Yaskawa INFORM job: -DEFRO-70-PRZYLACZE-70-NOWE.JBI

/JOB
//NAME -DEFRO-70-PRZYLACZE-70-NOWE
//POS
///NPOS 61,61,61,0,0,0
///TOOL 0
///POSTYPE PULSE
///PULSE
C00000=-281,-101163,-84214,3730,-80188,-1936
C00001=-283,-101162,-84213,3710,-80188,-1936
C00002=116617,-39062,-41553,1138,-40446,20
C00003=97332,10008,-65831,-77395,-56626,78097
C00004=97332,10036,-65835,-77406,-56622,78106
C00005=126597,-12792,-74683,9116,-14112,37031
C00006=129578,-9389,-72169,26197,-17561,29790
C00007=143171,23000,-49885,51799,-48783,19450
C00008=142289,27625,-43624,46606,-52109,19593
C00009=140707,34961,-33804,39360,-57405,19440
C00010=137188,46732,-18219,29241,-65914,18506
C00011=125601,64166,5444,7463,-78162,8461
C00012=120628,60223,2537,-370,-74792,3762
C00013=116260,63341,4618,-6746,-77452,-573
C00014=112604,59060,-1014,-13680,-74421,-638
C00015=105645,46181,-18056,-25918,-65595,-11662
C00016=96917,44348,-31091,-45677,-66308,-16214
C00017=100527,41964,-28031,-34606,-66372,-26006
C00018=106433,45775,-18486,-19914,-75527,-46558
C00019=110224,24520,-34980,-16270,-62186,-56055
C00020=117116,19907,-37131,-3644,-59039,-60958
C00021=117137,19542,-37273,-3641,-59137,-60967
C00022=117062,4461,-25894,-3265,-73866,-61376
C00023=116617,-39062,-41553,1138,-40446,20
C00024=97332,10008,-65831,-77395,-56626,78097
C00025=97332,10036,-65835,-77406,-56622,78106
C00026=126597,-12792,-74683,9116,-14112,37031
C00027=129578,-9389,-72169,26197,-17561,29790
C00028=143171,23000,-49885,51799,-48783,19450
C00029=142289,27625,-43624,46606,-52109,19593
C00030=140707,34961,-33804,39360,-57405,19440
C00031=137188,46732,-18219,29241,-65914,18506
C00032=125601,64166,5444,7463,-78162,8461
C00033=120628,60223,2537,-370,-74792,3762
C00034=116260,63341,4618,-6746,-77452,-573
C00035=112604,59060,-1014,-13680,-74421,-638
C00036=105645,46181,-18056,-25918,-65595,-11662
C00037=96917,44348,-31091,-45677,-66308,-16214
C00038=100527,41964,-28031,-34606,-66372,-26006
C00039=106433,45775,-18486,-19914,-75527,-46558
C00040=110224,24520,-34980,-16270,-62186,-56055
C00041=117116,19907,-37131,-3644,-59039,-60958
C00042=117137,19542,-37273,-3641,-59137,-60967
C00043=117062,4461,-25894,-3265,-73866,-61376
C00044=125074,-50101,-76658,51202,-17672,58606
C00045=125043,-41373,-84041,81327,-13668,44712
C00046=124776,-28424,-75745,87893,-13306,41755
C00047=124712,-28431,-75750,87904,-13268,41762
C00048=120787,-27884,-69765,25728,-8700,23794
C00049=115036,-25344,-64782,-26451,-15542,29683
C00050=119186,-28374,-69103,18427,-8940,-7851
C00051=122010,-28108,-68825,46224,-14319,-44839
C00052=116778,-25971,-65828,-246,-14948,-40490
C00053=118192,-23314,-61354,4708,-22161,-64875
C00054=115451,-27710,-69473,-21973,-12695,-70389
C00055=115429,-28374,-69925,-21919,-12759,-70410
C00056=115209,-37948,-70943,-16962,-16869,-72656
C00057=119279,-50675,-71302,9013,-26968,83196
C00058=116617,-39062,-41553,1138,-40446,20
C00059=-283,-101162,-84213,3710,-80188,-1936
C00060=-281,-101163,-84214,3730,-80188,-1936
BC00000=570125
BC00001=954451
BC00002=878037
BC00003=878036
BC00004=878036
BC00005=878037
BC00006=878037
BC00007=878037
BC00008=878037
BC00009=878037
BC00010=878037
BC00011=878037
BC00012=878036
BC00013=878037
BC00014=878037
BC00015=878037
BC00016=878037
BC00017=878037
BC00018=878037
BC00019=878037
BC00020=878037
BC00021=878037
BC00022=878037
BC00023=912351
BC00024=878036
BC00025=878036
BC00026=878037
BC00027=878037
BC00028=878037
BC00029=878037
BC00030=878037
BC00031=878037
BC00032=878037
BC00033=878036
BC00034=878037
BC00035=878037
BC00036=878037
BC00037=878037
BC00038=878037
BC00039=878037
BC00040=878037
BC00041=878037
BC00042=878037
BC00043=878037
BC00044=869720
BC00045=869720
BC00046=869720
BC00047=869720
BC00048=869721
BC00049=869721
BC00050=869721
BC00051=869721
BC00052=869721
BC00053=869721
BC00054=869721
BC00055=869721
BC00056=869721
BC00057=869720
BC00058=878037
BC00059=954451
BC00060=570125
EC00000=1163,0
EC00001=1166,0
EC00002=-1743,0
EC00003=-1746,0
EC00004=-1746,0
EC00005=-1743,0
EC00006=-1743,0
EC00007=-1743,0
EC00008=-1743,0
EC00009=-1743,0
EC00010=-1744,0
EC00011=-1744,0
EC00012=-1745,0
EC00013=-1744,0
EC00014=-1744,0
EC00015=-1744,0
EC00016=-1744,0
EC00017=-1744,0
EC00018=-1744,0
EC00019=-1744,0
EC00020=-1744,0
EC00021=-1744,0
EC00022=-1744,0
EC00023=-1743,0
EC00024=-1746,0
EC00025=-1746,0
EC00026=-1743,0
EC00027=-1743,0
EC00028=-1743,0
EC00029=-1743,0
EC00030=-1743,0
EC00031=-1744,0
EC00032=-1744,0
EC00033=-1745,0
EC00034=-1744,0
EC00035=-1744,0
EC00036=-1744,0
EC00037=-1744,0
EC00038=-1744,0
EC00039=-1744,0
EC00040=-1744,0
EC00041=-1744,0
EC00042=-1744,0
EC00043=-1744,0
EC00044=-85617,0
EC00045=-85617,0
EC00046=-85617,0
EC00047=-85617,0
EC00048=-85617,0
EC00049=-85617,0
EC00050=-85617,0
EC00051=-85617,0
EC00052=-85617,0
EC00053=-85617,0
EC00054=-85617,0
EC00055=-85617,0
EC00056=-85617,0
EC00057=-85617,0
EC00058=-1743,0
EC00059=1166,0
EC00060=1163,0
//INST
///DATE 2025/05/07 14:15
///ATTR SC,RW
///GROUP1 RB1,BS1
///GROUP2 ST1
NOP
MOVJ C00000 BC00000 VJ=80.00 DEC=20  +MOVJ EC00000 VJ=80.00
MOVJ C00001 BC00001 VJ=80.00 DEC=20  +MOVJ EC00001 VJ=0.78
MOVJ C00002 BC00002 VJ=80.00 DEC=20  +MOVJ EC00002 VJ=80.00
MOVJ C00003 BC00003 VJ=80.00 DEC=20  +MOVJ EC00003 VJ=2.00
TIMER T=0.50
MACRO1 MJ#(0) ARGF8
ARCON
WVON WEV#(21)
MOVC C00004 BC00004 V=5.0 DEC=20  +MOVJ EC00004 VJ=80.00
MOVC C00005 BC00005 V=5.0 DEC=20  +MOVJ EC00005 VJ=80.00
MOVC C00006 BC00006 V=5.0 DEC=20  +MOVJ EC00006 VJ=80.00
MOVL C00007 BC00007 V=5.0 DEC=20  +MOVJ EC00007 VJ=80.00
MOVL C00008 BC00008 V=7.5 DEC=20  +MOVJ EC00008 VJ=80.00
MOVL C00009 BC00009 V=5.0 DEC=20  +MOVJ EC00009 VJ=0.78
MOVC C00010 BC00010 V=5.0 DEC=20  +MOVJ EC00010 VJ=80.00
MOVC C00011 BC00011 V=5.0 DEC=20  +MOVJ EC00011 VJ=80.00
WVON WEV#(22)
MOVC C00012 BC00012 V=5.0 DEC=20  +MOVJ EC00012 VJ=80.00
MOVC C00013 BC00013 V=5.0 DEC=20  +MOVJ EC00013 VJ=80.00
WVON WEV#(23)
MOVC C00014 BC00014 V=5.0 DEC=20  +MOVJ EC00014 VJ=80.00
MOVC C00015 BC00015 V=5.0 DEC=20  +MOVJ EC00015 VJ=80.00
MOVL C00016 BC00016 V=5.0 DEC=20  +MOVJ EC00016 VJ=80.00
MOVL C00017 BC00017 V=7.5 DEC=20  +MOVJ EC00017 VJ=80.00
WVON WEV#(21)
MOVC C00018 BC00018 V=6.7 DEC=20  +MOVJ EC00018 VJ=80.00
MOVL C00019 BC00019 V=5.0 DEC=20  +MOVJ EC00019 VJ=80.00
MOVL C00020 BC00020 V=5.0 DEC=20  +MOVJ EC00020 VJ=80.00
MOVC C00021 BC00021 V=5.0 DEC=20  +MOVJ EC00021 VJ=80.00
ARCOF
WVOF
MOVJ C00022 BC00022 VJ=80.00 DEC=20  +MOVJ EC00022 VJ=80.00
MOVJ C00023 BC00023 VJ=80.00 DEC=20  +MOVJ EC00023 VJ=80.00
MOVJ C00024 BC00024 VJ=80.00 DEC=20  +MOVJ EC00024 VJ=2.00
TIMER T=0.50
MACRO1 MJ#(0) ARGF8
ARCON
WVON WEV#(21)
MOVC C00025 BC00025 V=5.0 DEC=20  +MOVJ EC00025 VJ=80.00
MOVC C00026 BC00026 V=5.0 DEC=20  +MOVJ EC00026 VJ=80.00
MOVC C00027 BC00027 V=5.0 DEC=20  +MOVJ EC00027 VJ=80.00
MOVL C00028 BC00028 V=5.0 DEC=20  +MOVJ EC00028 VJ=80.00
MOVL C00029 BC00029 V=7.5 DEC=20  +MOVJ EC00029 VJ=80.00
MOVL C00030 BC00030 V=5.0 DEC=20  +MOVJ EC00030 VJ=0.78
MOVC C00031 BC00031 V=5.0 DEC=20  +MOVJ EC00031 VJ=80.00
MOVC C00032 BC00032 V=5.0 DEC=20  +MOVJ EC00032 VJ=80.00
WVON WEV#(22)
MOVC C00033 BC00033 V=5.0 DEC=20  +MOVJ EC00033 VJ=80.00
MOVC C00034 BC00034 V=5.0 DEC=20  +MOVJ EC00034 VJ=80.00
WVON WEV#(23)
MOVC C00035 BC00035 V=5.0 DEC=20  +MOVJ EC00035 VJ=80.00
MOVC C00036 BC00036 V=5.0 DEC=20  +MOVJ EC00036 VJ=80.00
MOVL C00037 BC00037 V=5.0 DEC=20  +MOVJ EC00037 VJ=80.00
MOVL C00038 BC00038 V=7.5 DEC=20  +MOVJ EC00038 VJ=80.00
WVON WEV#(21)
MOVC C00039 BC00039 V=6.7 DEC=20  +MOVJ EC00039 VJ=80.00
MOVL C00040 BC00040 V=5.0 DEC=20  +MOVJ EC00040 VJ=80.00
MOVL C00041 BC00041 V=5.0 DEC=20  +MOVJ EC00041 VJ=80.00
MOVC C00042 BC00042 V=5.0 DEC=20  +MOVJ EC00042 VJ=80.00
ARCOF
WVOF
MOVJ C00043 BC00043 VJ=80.00 DEC=20  +MOVJ EC00043 VJ=80.00
MOVJ C00044 BC00044 VJ=80.00 DEC=20  +MOVJ EC00044 VJ=80.00
MOVJ C00045 BC00045 VJ=80.00 DEC=20  +MOVJ EC00045 VJ=80.00
MOVJ C00046 BC00046 VJ=80.00 DEC=20  +MOVJ EC00046 VJ=80.00
TIMER T=0.50
MACRO1 MJ#(0) ARGF4
ARCON
MOVC C00047 BC00047 V=5.0 DEC=20  +MOVJ EC00047 VJ=80.00
MOVC C00048 BC00048 V=5.0 DEC=20  +MOVJ EC00048 VJ=80.00
MOVC C00049 BC00049 V=5.0 DEC=20  +MOVJ EC00049 VJ=80.00
MOVC C00050 BC00050 V=5.0 DEC=20  +MOVJ EC00050 VJ=80.00
MOVC C00051 BC00051 V=5.0 DEC=20  +MOVJ EC00051 VJ=80.00
MOVC C00052 BC00052 V=5.0 DEC=20  +MOVJ EC00052 VJ=80.00
MOVC C00053 BC00053 V=5.0 DEC=20  +MOVJ EC00053 VJ=80.00
MOVC C00054 BC00054 V=5.0 DEC=20  +MOVJ EC00054 VJ=80.00
MOVJ C00055 BC00055 VJ=2.00 DEC=20  +MOVJ EC00055 VJ=80.00
ARCOF
MOVJ C00056 BC00056 VJ=80.00 DEC=20  +MOVJ EC00056 VJ=80.00
MOVJ C00057 BC00057 VJ=80.00 DEC=20  +MOVJ EC00057 VJ=80.00
MOVJ C00058 BC00058 VJ=80.00 DEC=20  +MOVJ EC00058 VJ=80.00
MOVJ C00059 BC00059 VJ=80.00 DEC=20  +MOVJ EC00059 VJ=80.00
MOVJ C00060 BC00060 VJ=80.00 DEC=20  +MOVJ EC00060 VJ=80.00
END
